// TIA Portal V19 export
DATA_BLOCK "RVL"   // DB3
{ S7_Optimized_Access := 'TRUE' }
// stored: MemoryReserve 100
   VAR
      ConveyorVelocity : Array[0..10] of Real;   // mmps
   END_VAR
BEGIN
   ConveyorVelocity[0] := 500.0;
   ConveyorVelocity[1] := 700.0;
   ConveyorVelocity[2] := 500.0;
   ConveyorVelocity[3] := 50.0;
   ConveyorVelocity[4..5] := 500.0;
   ConveyorVelocity[6..10] := 50.0;
END_DATA_BLOCK
